// TIA Portal V19 export
// export: Created 2026-10-15T09:44:25.2469114Z, ExportSetting WithDefaults, DisplayName Totally Integrated Automation Portal, DisplayVersion V19, DisplayName TIA Portal Openness, DisplayVersion V19, DisplayName TIA Portal Version Control Interface, DisplayVersion V19, DisplayName STEP 7 Professional, DisplayVersion V19, DisplayName STEP 7 Safety, DisplayVersion V19, DisplayName WinCC Basic/Comfort/Advanced, DisplayVersion V19, DisplayName WinCC Unified, DisplayVersion V19
FUNCTION "ROLL_ReadInputs" : Void   // FC36, SCL
{ S7_Optimized_Access := 'TRUE' }
VERSION : 0.1
// stored: AutoNumber true, IsIECCheckEnabled false, SetENOAutomatically false, UDAEnableTagReadback false
   VAR_TEMP
      "b" : Int;
      bit : Int;
   END_VAR
BEGIN

   // Confirmed four-station profile: absent optional inputs are zero.
   FOR #b := 119 TO 125 DO
       FOR #bit := 0 TO 7 DO
           "ROLL_IO".Input[#b, #bit] := FALSE;
       END_FOR;
   END_FOR;
   IF "ROLL_IO".PhysicalIoConfigured AND NOT "ROLL_IO".Simulation THEN
       "ROLL_IO".Input[0, 0] := "Tag__639276542175325643";
       "ROLL_IO".Input[0, 1] := "Tag__639276542176642122";
       "ROLL_IO".Input[0, 2] := "Tag__639276542176711934";
       "ROLL_IO".Input[0, 3] := "Tag__639276542176781759";
       "ROLL_IO".Input[0, 4] := "Tag__639276542176841598";
       "ROLL_IO".Input[0, 5] := "Tag__639276542176901438";
       "ROLL_IO".Input[0, 6] := "Tag__639276542176961268";
       "ROLL_IO".Input[0, 7] := "Tag__639276542177021200";
       "ROLL_IO".Input[1, 0] := "Tag__639276542177080956";
       "ROLL_IO".Input[1, 1] := "Tag__639276542177140787";
       "ROLL_IO".Input[1, 2] := "Tag__639276542177200628";
       "ROLL_IO".Input[1, 3] := "Tag__639276542177260475";
       "ROLL_IO".Input[1, 4] := "Tag__639276542177320320";
       "ROLL_IO".Input[1, 5] := "Tag__639276542177370179";
       "ROLL_IO".Input[1, 6] := "Tag__639276542177430014";
       "ROLL_IO".Input[1, 7] := "Tag__639276542177499830";
       "ROLL_IO".Input[2, 0] := "Tag__639276542177559666";
       "ROLL_IO".Input[2, 1] := "Tag__639276542177609533";
       "ROLL_IO".Input[2, 2] := "Tag__639276542177669373";
       "ROLL_IO".Input[2, 3] := "Tag__639276542177729387";
       "ROLL_IO".Input[2, 4] := "Tag__639276542177789061";
       "ROLL_IO".Input[2, 5] := "Tag__639276542177848893";
       "ROLL_IO".Input[2, 6] := "Tag__639276542177898771";
       "ROLL_IO".Input[2, 7] := "Tag__639276542177958599";
       "ROLL_IO".Input[3, 0] := "Tag__639276542178018439";
       "ROLL_IO".Input[3, 1] := "Tag__639276542178078280";
       "ROLL_IO".Input[3, 2] := "Tag__639276542178138119";
       "ROLL_IO".Input[3, 3] := "Tag__639276542178197968";
       "ROLL_IO".Input[3, 4] := "Tag__639276542178257802";
       "ROLL_IO".Input[3, 5] := "Tag__639276542178317647";
       "ROLL_IO".Input[3, 6] := "Tag__639276542178377487";
       "ROLL_IO".Input[3, 7] := "Tag__639276542178427358";
       "ROLL_IO".Input[4, 0] := "Tag__639276542178487269";
       "ROLL_IO".Input[4, 1] := "Tag__639276542178547298";
       "ROLL_IO".Input[4, 2] := "Tag__639276542178607019";
       "ROLL_IO".Input[4, 3] := "Tag__639276542178666705";
       "ROLL_IO".Input[4, 4] := "Tag__639276542178726546";
       "ROLL_IO".Input[4, 5] := "Tag__639276542178776412";
       "ROLL_IO".Input[4, 6] := "Tag__639276542178836252";
       "ROLL_IO".Input[4, 7] := "Tag__639276542178896091";
       "ROLL_IO".Input[5, 0] := "Tag__639276542178955944";
       "ROLL_IO".Input[5, 1] := "Tag__639276542179015839";
       "ROLL_IO".Input[5, 2] := "Tag__639276542179085589";
       "ROLL_IO".Input[5, 3] := "Tag__639276542179135453";
       "ROLL_IO".Input[5, 4] := "Tag__639276542179195720";
       "ROLL_IO".Input[5, 5] := "Tag__639276542179255406";
       "ROLL_IO".Input[5, 6] := "Tag__639276542179314975";
       "ROLL_IO".Input[5, 7] := "Tag__639276542179384784";
       "ROLL_IO".Input[6, 0] := "Tag__639276542179434654";
       "ROLL_IO".Input[6, 1] := "Tag__639276542179494489";
       "ROLL_IO".Input[6, 2] := "Tag__639276542179554331";
       "ROLL_IO".Input[6, 3] := "Tag__639276542179614187";
       "ROLL_IO".Input[6, 4] := "Tag__639276542179674010";
       "ROLL_IO".Input[6, 5] := "Tag__639276542179723877";
       "ROLL_IO".Input[6, 6] := "Tag__639276542179783716";
       "ROLL_IO".Input[6, 7] := "Tag__639276542179843556";
       "ROLL_IO".Input[7, 0] := "Tag__639276542179903396";
       "ROLL_IO".Input[7, 1] := "Tag__639276542179963535";
       "ROLL_IO".Input[7, 2] := "Tag__639276542180023076";
       "ROLL_IO".Input[7, 3] := "Tag__639276542180082916";
       "ROLL_IO".Input[7, 4] := "Tag__639276542180142913";
       "ROLL_IO".Input[7, 5] := "Tag__639276542180202595";
       "ROLL_IO".Input[7, 6] := "Tag__639276542180262436";
       "ROLL_IO".Input[7, 7] := "Tag__639276542180322276";
       "ROLL_IO".Input[8, 0] := "Tag__639276542180382124";
       "ROLL_IO".Input[8, 1] := "Tag__639276542180441967";
       "ROLL_IO".Input[8, 2] := "Tag__639276542180501796";
       "ROLL_IO".Input[8, 3] := "Tag__639276542180561959";
       "ROLL_IO".Input[8, 4] := "Tag__639276542180621475";
       "ROLL_IO".Input[8, 5] := "Tag__639276542180681324";
       "ROLL_IO".Input[8, 6] := "Tag__639276542180741155";
       "ROLL_IO".Input[8, 7] := "Tag__639276542180801004";
       "ROLL_IO".Input[9, 0] := "Tag__639276542180860838";
       "ROLL_IO".Input[9, 1] := "Tag__639276542180920674";
       "ROLL_IO".Input[9, 2] := "Tag__639276542180980515";
       "ROLL_IO".Input[9, 3] := "Tag__639276542181040355";
       "ROLL_IO".Input[9, 4] := "Tag__639276542181100204";
       "ROLL_IO".Input[9, 5] := "Tag__639276542181160040";
       "ROLL_IO".Input[9, 6] := "Tag__639276542181219884";
       "ROLL_IO".Input[9, 7] := "Tag__639276542181289692";
       "ROLL_IO".Input[10, 0] := "Tag__639276542181349527";
       "ROLL_IO".Input[10, 1] := "Tag__639276542181429316";
       "ROLL_IO".Input[10, 2] := "Tag__639276542181489163";
       "ROLL_IO".Input[10, 3] := "Tag__639276542181548993";
       "ROLL_IO".Input[10, 4] := "Tag__639276542181608833";
       "ROLL_IO".Input[10, 5] := "Tag__639276542181668673";
       "ROLL_IO".Input[10, 6] := "Tag__639276542181728514";
       "ROLL_IO".Input[10, 7] := "Tag__639276542181778645";
       "ROLL_IO".Input[11, 0] := "Tag__639276542181848196";
       "ROLL_IO".Input[11, 1] := "Tag__639276542181937992";
       "ROLL_IO".Input[11, 2] := "Tag__639276542182007903";
       "ROLL_IO".Input[11, 3] := "Tag__639276542182097533";
       "ROLL_IO".Input[11, 4] := "Tag__639276542182167640";
       "ROLL_IO".Input[11, 5] := "Tag__639276542182237171";
       "ROLL_IO".Input[11, 6] := "Tag__639276542182316955";
       "ROLL_IO".Input[11, 7] := "Tag__639276542182396730";
       "ROLL_IO".Input[12, 0] := "Tag__639276542182476554";
       "ROLL_IO".Input[12, 1] := "Tag__639276542182566280";
       "ROLL_IO".Input[12, 2] := "Tag__639276542182636090";
       "ROLL_IO".Input[12, 3] := "Tag__639276542182715877";
       "ROLL_IO".Input[12, 4] := "Tag__639276542182795660";
       "ROLL_IO".Input[12, 5] := "Tag__639276542182855499";
       "ROLL_IO".Input[12, 6] := "Tag__639276542182915345";
       "ROLL_IO".Input[12, 7] := "Tag__639276542182975191";
       "ROLL_IO".Input[13, 0] := "Tag__639276542183035019";
       "ROLL_IO".Input[13, 1] := "Tag__639276542183094859";
       "ROLL_IO".Input[13, 2] := "Tag__639276542183154975";
       "ROLL_IO".Input[13, 3] := "Tag__639276542183214549";
       "ROLL_IO".Input[13, 4] := "Tag__639276542183274379";
       "ROLL_IO".Input[13, 5] := "Tag__639276542183334218";
       "ROLL_IO".Input[13, 6] := "Tag__639276542183394068";
       "ROLL_IO".Input[13, 7] := "Tag__639276542183453907";
       "ROLL_IO".Input[14, 0] := "Tag__639276542183523712";
       "ROLL_IO".Input[14, 1] := "Tag__639276542183583551";
       "ROLL_IO".Input[14, 2] := "Tag__639276542183643721";
       "ROLL_IO".Input[14, 3] := "Tag__639276542183703360";
       "ROLL_IO".Input[14, 4] := "Tag__639276542183763071";
       "ROLL_IO".Input[14, 5] := "Tag__639276542183822911";
       "ROLL_IO".Input[14, 6] := "Tag__639276542183883174";
       "ROLL_IO".Input[14, 7] := "Tag__639276542183942603";
       "ROLL_IO".Input[15, 0] := "Tag__639276542184002441";
       "ROLL_IO".Input[15, 1] := "Tag__639276542184072244";
       "ROLL_IO".Input[15, 2] := "Tag__639276542184132093";
       "ROLL_IO".Input[15, 3] := "Tag__639276542184181958";
       "ROLL_IO".Input[15, 4] := "Tag__639276542184241948";
       "ROLL_IO".Input[15, 5] := "Tag__639276542184301629";
       "ROLL_IO".Input[15, 6] := "Tag__639276542184361470";
       "ROLL_IO".Input[15, 7] := "Tag__639276542184421310";
   END_IF;
END_FUNCTION
